// TIA Portal V21 export
// export: Created 2026-11-10T07:35:22.3630755Z, ExportSetting WithDefaults, DisplayName Totally Integrated Automation Portal, DisplayVersion V21 Update 3, DisplayName STEP 7 Professional, DisplayVersion V21 Update 3, DisplayName STEP 7 Safety, DisplayVersion V21, DisplayName Tech WebApplication, DisplayVersion V21, DisplayName WinCC Basic/Comfort/Advanced, DisplayVersion V21 Update 3, DisplayName WinCC Unified, DisplayVersion V21 Update 3
FUNCTION_BLOCK "FB_Lad_ex151"   // FB55, LAD
{ S7_Optimized_Access := 'TRUE' }
VERSION : 0.1
// stored: AutoNumber true, IsIECCheckEnabled false, IsRetainMemResEnabled false, MemoryReserve 100, SetENOAutomatically false, UDAEnableTagReadback false
   VAR_INPUT
      v_req : Bool;
      v_db_number : UInt;
   END_VAR
   VAR_OUTPUT
      v_ret_val : Int;
      v_busy : Bool;
   END_VAR
BEGIN

REGION Network 1: DELETE_DB - Delete data block
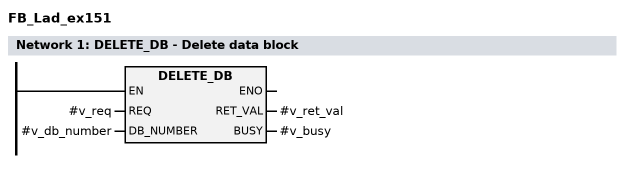
   RUNG wire#powerrail
      DELETE_DB(REQ := #v_req, DB_NUMBER := #v_db_number, Ret_Val => #v_ret_val, BUSY => #v_busy)
   END_RUNG
   // the same network as SCL:
   #v_ret_val := DELETE_DB(REQ := #v_req, DB_NUMBER := #v_db_number, BUSY => #v_busy);
END_REGION
END_FUNCTION_BLOCK
